Fanuc KAREL source: kx00005.KL

-- PROVISIONAL review KL for V940-1; original PC SHA256 501246f717d869685a48993f7bbf3493dcb52a4530bc86edf102abf405565ad8
-- Incomplete behavior may be omitted. Consult companion uncertainty JSON. Do not deploy.
PROGRAM KX00005
%NOLOCKGROUP
VAR
  I : INTEGER
  J : INTEGER
  B : BOOLEAN
  F : FILE
  S : STRING[80]
-- UNRESOLVED_DECL P type=000102
BEGIN
  -- V9_ZERO_TABLE_METADATA_HINT layout=0001; no indexed target words; source/name/runtime held
  -- UNRESOLVED_PC offsets 5-32; opcodes 22,3F,3F,3D
  -- UNRESOLVED_PC offsets 37-44; opcodes 22,A3
  -- UNRESOLVED_PC offsets 49-56; opcodes 22,39
  -- UNRESOLVED_PC offsets 61-65; opcodes 7F
END KX00005
